FUNCTION_BLOCK FB_LightTests EXTENDS TcUnit.FB_TestSuite
VAR
END_VAR

ToggleTurnsLightOn();
SecondToggleTurnsLightOff();
NoToggleKeepsCurrentState();
HeldToggleDoesNotRetrigger();
ToggleRearminAfterRelease();
SetRequestsForceState();
ToggleWinsOverSetRequest();
IndependentLightsKeepIndependentState();

METHOD PRIVATE HeldToggleDoesNotRetrigger
VAR
    fbLight : FB_Light;
END_VAR
TEST('Held toggle does not retrigger');
fbLight.bToggle := TRUE;
fbLight();
fbLight();
AssertTrue(Condition := fbLight.bOn, Message := 'Held toggle should only turn the light on once');
TEST_FINISHED();
END_METHOD

METHOD PRIVATE ToggleRearminAfterRelease
VAR
    fbLight : FB_Light;
END_VAR
TEST('Toggle rearms after release');
fbLight.bToggle := TRUE;
fbLight();
fbLight.bToggle := FALSE;
fbLight();
fbLight.bToggle := TRUE;
fbLight();
AssertFalse(Condition := fbLight.bOn, Message := 'A new rising edge should turn the light off');
TEST_FINISHED();
END_METHOD

METHOD PRIVATE SetRequestsForceState
VAR
    fbLight : FB_Light;
END_VAR
TEST('Set requests force state');
fbLight.bSetValid := TRUE;
fbLight.bSetOn := TRUE;
fbLight();
AssertTrue(Condition := fbLight.bOn, Message := 'Valid ON request should turn light on');
fbLight.bSetOn := FALSE;
fbLight();
AssertFalse(Condition := fbLight.bOn, Message := 'Valid OFF request should turn light off');
fbLight.bSetValid := FALSE;
fbLight.bSetOn := TRUE;
fbLight();
AssertFalse(Condition := fbLight.bOn, Message := 'Invalid set request should be ignored');
TEST_FINISHED();
END_METHOD

METHOD PRIVATE ToggleWinsOverSetRequest
VAR
    fbLight : FB_Light;
END_VAR
TEST('Toggle wins over set request');
fbLight.bToggle := TRUE;
fbLight.bSetValid := TRUE;
fbLight.bSetOn := FALSE;
fbLight();
AssertTrue(Condition := fbLight.bOn, Message := 'Toggle should win over simultaneous set OFF request');
TEST_FINISHED();
END_METHOD

METHOD PRIVATE IndependentLightsKeepIndependentState
VAR
    fbLight1 : FB_Light;
    fbLight2 : FB_Light;
END_VAR
TEST('Independent lights keep independent state');
fbLight1.bToggle := TRUE;
fbLight1();
fbLight2();
AssertTrue(Condition := fbLight1.bOn, Message := 'First light should be on');
AssertFalse(Condition := fbLight2.bOn, Message := 'Second light should remain off');
TEST_FINISHED();
END_METHOD

METHOD PRIVATE NoToggleKeepsCurrentState
VAR
    fbLight : FB_Light;
END_VAR
TEST('No toggle keeps current state');
fbLight();
AssertFalse(Condition := fbLight.bOn, Message := 'Light should remain OFF without toggle');
TEST_FINISHED();
END_METHOD

METHOD PRIVATE SecondToggleTurnsLightOff
VAR
    fbLight : FB_Light;
END_VAR
TEST('Second toggle turns light off');
fbLight.bToggle := TRUE;
fbLight();
fbLight.bToggle := FALSE;
fbLight();
fbLight.bToggle := TRUE;
fbLight();
AssertFalse(Condition := fbLight.bOn, Message := 'Second toggle should turn light off');
TEST_FINISHED();
END_METHOD

METHOD PRIVATE ToggleTurnsLightOn
VAR
    fbLight : FB_Light;
END_VAR
TEST('Toggle turns light on');
fbLight.bToggle := TRUE;
fbLight();
AssertTrue(Condition := fbLight.bOn, Message := 'Toggle should turn light on');
TEST_FINISHED();
END_METHOD

END_FUNCTION_BLOCK

(* stored: Version 1.1.0.1
   POU FB_LightTests: Id {c5856838-1d6b-4b34-b900-07483f8bff5f}, SpecialFunc None
   Method HeldToggleDoesNotRetrigger: Id {371fc64a-d964-4d52-8a5d-8e401ded155e}
   Method ToggleRearminAfterRelease: Id {24b4f532-0e77-41d4-a348-8c3d6b490c41}
   Method SetRequestsForceState: Id {947ee51d-6209-4674-b58d-0491d1856139}
   Method ToggleWinsOverSetRequest: Id {87a1a087-3516-4a42-a79b-aa437ee90c5f}
   Method IndependentLightsKeepIndependentState: Id {62fa420d-cd87-47fc-a5c8-970cf7f5848f}
   Method NoToggleKeepsCurrentState: Id {3f7c2d53-b707-4069-ae01-d00505e72865}
   Method SecondToggleTurnsLightOff: Id {8b0859e6-a360-4010-b172-3025a975b5c7}
   Method ToggleTurnsLightOn: Id {0219653a-ebc7-4f44-b312-192b3fedd447} *)
